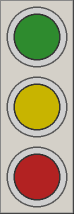
VISUALIZATION Vis_LightTower  // 74x214
    Rectangle (0,0 74x214), colour toggle: prg_LightTower.qBuzzer
    Lamp1 (2,2 70x70), variable: prg_LightTower.qLedGreen, style: Lamp-Lamp1-Green
    Lamp1 (2,72 70x70), variable: prg_LightTower.qLedYellow, style: Lamp-Lamp1-Yellow
    Lamp1 (2,142 70x70), variable: prg_LightTower.qLedRed, style: Lamp-Lamp1-Red
END_VISUALIZATION

(* stored: Version 1.1.0.1, ProductVersion 3.1.4024.13
   Visu Vis_LightTower: Id {c021278b-318c-482e-8d29-2836dfb07464} *)
